(* IEC 61131-3 sources: nautilus/examples/it-cluster/lib, 2 files *)

(* ---- server.st ---- *)
(* The server half of the plant: fault inputs, a first-order thermal model,
   and how a server's parts respond. Same rules as lib/switch.st: a fault
   is an input, the recording is the baseline, faults compose, clearing a
   fault lets the recording show through again.

   The thermal model is deliberately small, and every number that shapes it
   is a named constant below, to tune against what a real box does:

     load rise    = KLoad * (CpuLoad - RecLoadPct)
     rise target  = load rise
                  + KFanFrac * failed fans * (CPU over inlet + load rise)
                  - KBoostCool * (FanBoost - 1)         the others ramping
     each sensor  = recorded + Weight * rise + room offset, approached
                    with time constant TauS (first order), so a failure
                    makes temperatures CLIMB rather than jump
     fan boost    = 1 + KBoost * (CPU rise now), capped at MaxBoost: the
                    BMC's fan curve answering the temperature it reads

   Where the numbers come from (the node is a Supermicro 1U with one
   Xeon 6505P: 150 W TDP, 97 °C DTS max; its BMC calls 102 °C critical):
     WPerPct   150 W TDP over an idle package of about 35 W, across 90 %
               of load: about 1.3 W per %
     KLoad     that power through a 1U heatsink at about 0.3 °C/W:
               about 0.35 °C per %
     KFanFrac  one of six fans gone costs the heatsink about a fifth of its
               airflow; its thermal resistance, and so the CPU's rise over
               the inlet, grows by about as much: small at idle, large
               under load, which is how a lost fan really behaves
     TauS      a 1U heatsink under forced air settles in about a minute
               (vendors give 60 s to swap a fan before cooling is lost)
     CapC      the CPU throttles near its limit rather than running away:
               held a little past the BMC's critical, so the alarm trips *)

TYPE
  SimServer : STRUCT
    Dark     : BOOL; (* the BMC stops answering: Online false *)
    PowerOff : BOOL; (* host off: standby power, fans stop, temps fall to inlet, host links drop; the BMC stays up *)
    CpuLoad  : REAL; (* % busy, 0 = as recorded (the recording is a quiet cluster, about RecLoadPct) *)
  END_STRUCT;
  SimFan : STRUCT
    Fail : BOOL; (* stopped: RPM 0, Fault; the other fans ramp, temperatures rise *)
  END_STRUCT;
  SimPSU : STRUCT
    InputLost : BOOL; (* line cord out: InputOk false, output 0, the other PSU carries the load *)
    Fail      : BOOL; (* the supply itself fails: Fault, output 0 *)
  END_STRUCT;
  SimDrive : STRUCT
    Pulled  : BOOL; (* out of its bay: Present false *)
    Failing : BOOL; (* SMART predicts failure: PredictedFailure, health Warning *)
  END_STRUCT;
  SimNetPort : STRUCT
    Down : BOOL; (* the port loses link: both ends of its cable go down *)
  END_STRUCT;
  SimCable : STRUCT
    Pulled : BOOL; (* the cable itself: both ends down *)
  END_STRUCT;
  SimRoom : STRUCT
    InletDeltaC : REAL; (* the room runs hot: every server's inlet, and everything behind it, rises *)
  END_STRUCT;
END_TYPE

FUNCTION_BLOCK ServerPlant
(* The chassis: power, CPU busy, and the thermal model's rise. Its outputs
   drive the fans, sensors and PSUs of the same server. *)
VAR_INPUT
  Rec        : Server;
  F          : SimServer;
  Room       : SimRoom;
  FansFailed : DINT;
  CpuRiseNow : REAL; (* the CPU sensor's current rise over the recording, for the fan curve *)
  CpuOverInlet : REAL := 35.0; (* the recorded CPU temperature above the recorded inlet *)
  Live       : BOOL;
  Unpowered  : BOOL; (* every supply down (plant.st): no standby power either *)
END_VAR
VAR_IN_OUT
  P : Server;
END_VAR
VAR_OUTPUT
  RiseTarget : REAL; (* °C the CPU heads for above the recording *)
  FanBoost   : REAL; (* the fans' speed factor *)
  Off        : BOOL;
  Dead       : BOOL; (* no power at all: the host off and the BMC with it *)
  LoadW      : REAL; (* the power the PSUs deliver *)
END_VAR
VAR
  B        : Server;
  Init     : BOOL;
  LoadRise : REAL;
END_VAR
VAR CONSTANT
  RecLoadPct : REAL := 10.0;  (* the recording's CPU busy: an idle cluster *)
  KLoad      : REAL := 0.35;  (* °C per % of extra load *)
  KFanFrac   : REAL := 0.2;   (* per failed fan: the share by which the CPU's rise over the inlet grows *)
  KBoost     : REAL := 0.03;  (* fan speed-up per °C of CPU rise *)
  MaxBoost   : REAL := 1.6;   (* fans at their ceiling *)
  KBoostCool : REAL := 10.0;  (* °C the ramped fans take back at full boost - 1 *)
  WPerPct    : REAL := 1.3;   (* W per % of extra load *)
  StandbyW   : REAL := 12.0;  (* host off, BMC on *)
END_VAR
IF NOT Init THEN
  B := P;
  Init := TRUE;
END_IF;
IF Live THEN
  B.PowerOn := Rec.PowerOn;
  B.PowerW := Rec.PowerW;
  B.InletTempC := Rec.InletTempC;
  B.MaxTempC := Rec.MaxTempC;
END_IF;
Dead := Unpowered;
Off := F.PowerOff OR NOT B.PowerOn OR Dead;
P.Online := NOT (F.Dark OR Dead);
P.PowerOn := NOT Off;
FanBoost := LIMIT(1.0, 1.0 + KBoost * MAX(CpuRiseNow, 0.0), MaxBoost);
IF Off THEN
  RiseTarget := 0.0;
  LoadW := SEL(Dead, StandbyW, 0.0);
  P.CpuPct := 0.0;
ELSE
  LoadRise := 0.0;
  IF F.CpuLoad > 0.0 THEN
    LoadRise := KLoad * (F.CpuLoad - RecLoadPct);
  END_IF;
  RiseTarget := LoadRise + KFanFrac * INT_TO_REAL(FansFailed) * MAX(CpuOverInlet + LoadRise, 0.0)
    - KBoostCool * (FanBoost - 1.0);
  IF F.CpuLoad > 0.0 THEN
    LoadW := B.PowerW + WPerPct * (F.CpuLoad - RecLoadPct);
    P.CpuPct := F.CpuLoad;
  ELSE
    LoadW := B.PowerW;
    P.CpuPct := RecLoadPct;
  END_IF;
END_IF;
P.PowerW := LoadW;
P.InletTempC := B.InletTempC + Room.InletDeltaC;
END_FUNCTION_BLOCK

FUNCTION_BLOCK TempPlant
(* One temperature sensor: its recording, plus Weight x the server's rise,
   plus the room; approached with TauS. Off, it cools to the inlet. *)
VAR_INPUT
  Rec        : TempSensor;
  RiseTarget : REAL;
  Weight     : REAL; (* 1 for the CPU, less for what sits further from it, 0 for the inlet *)
  RoomC      : REAL;
  InletC     : REAL; (* where it cools to, host off *)
  Off        : BOOL;
  Dt         : REAL;
  Live       : BOOL;
  CapC       : REAL := 110.0; (* where the part throttles or trips; the CPU's is lower *)
END_VAR
VAR_IN_OUT
  P : TempSensor;
END_VAR
VAR_OUTPUT
  Rise : REAL; (* now, over the recording *)
  Base : REAL; (* the recording (or snapshot) *)
END_VAR
VAR
  B     : TempSensor;
  Init  : BOOL;
  State : REAL; (* the sensor's own lagged offset from the recording *)
  Goal  : REAL;
END_VAR
VAR CONSTANT
  TauS    : REAL := 60.0;  (* heating and cooling time constant *)
  OffTauS : REAL := 300.0; (* cooling to the inlet, host off *)
END_VAR
IF NOT Init THEN
  B := P;
  Init := TRUE;
END_IF;
IF Live THEN
  B.Value := Rec.Value;
END_IF;
IF Off THEN
  Goal := InletC - B.Value;
  State := State + (Goal - State) * MIN(Dt / OffTauS, 1.0);
ELSE
  Goal := Weight * RiseTarget + RoomC;
  State := State + (Goal - State) * MIN(Dt / TauS, 1.0);
END_IF;
P.Value := MIN(B.Value + State, CapC);
Rise := P.Value - B.Value;
Base := B.Value;
P.High := P.HighSP > 0.0 AND P.Value >= P.HighSP;
P.HighHigh := P.HighHighSP > 0.0 AND P.Value >= P.HighHighSP;
END_FUNCTION_BLOCK

FUNCTION_BLOCK FanPlant
VAR_INPUT
  Rec   : Fan;
  F     : SimFan;
  Boost : REAL;
  Off   : BOOL;
  Live  : BOOL;
END_VAR
VAR_IN_OUT
  P : Fan;
END_VAR
VAR
  B    : Fan;
  Init : BOOL;
END_VAR
VAR CONSTANT
  MaxRPM : REAL := 16000.0;
END_VAR
IF NOT Init THEN
  B := P;
  Init := TRUE;
END_IF;
IF Live THEN
  B.RPM := Rec.RPM;
END_IF;
IF F.Fail OR Off THEN
  P.RPM := 0.0;
ELSE
  P.RPM := MIN(B.RPM * Boost, MaxRPM);
END_IF;
P.Fault := F.Fail;
END_FUNCTION_BLOCK

FUNCTION_BLOCK PsuPair
(* Two supplies sharing a load: each carries its recorded share while both
   are up; one lost, the other carries it all and the server stays up; both
   lost, neither carries anything (the server is Unpowered, plant.st). *)
VAR_INPUT
  Rec1, Rec2 : PSU;
  F1, F2     : SimPSU;
  LoadW      : REAL;
  Live       : BOOL;
END_VAR
VAR_IN_OUT
  P1, P2 : PSU;
END_VAR
VAR
  B1, B2 : PSU;
  Init   : BOOL;
  Up1, Up2 : BOOL;
  Share1 : REAL;
END_VAR
IF NOT Init THEN
  B1 := P1;
  B2 := P2;
  Init := TRUE;
END_IF;
IF Live THEN
  B1.InputV := Rec1.InputV;
  B1.OutputW := Rec1.OutputW;
  B2.InputV := Rec2.InputV;
  B2.OutputW := Rec2.OutputW;
END_IF;
Up1 := NOT (F1.InputLost OR F1.Fail);
Up2 := NOT (F2.InputLost OR F2.Fail);
Share1 := 0.5;
IF B1.OutputW + B2.OutputW > 0.0 THEN
  Share1 := B1.OutputW / (B1.OutputW + B2.OutputW);
END_IF;
IF NOT Up2 THEN
  Share1 := 1.0;
ELSIF NOT Up1 THEN
  Share1 := 0.0;
END_IF;
P1.OutputW := LoadW * Share1;
P2.OutputW := LoadW * (1.0 - Share1);
IF NOT (Up1 OR Up2) THEN
  P1.OutputW := 0.0;
  P2.OutputW := 0.0;
END_IF;
P1.InputOk := NOT F1.InputLost;
P2.InputOk := NOT F2.InputLost;
P1.InputV := SEL(F1.InputLost, B1.InputV, 0.0);
P2.InputV := SEL(F2.InputLost, B2.InputV, 0.0);
(* a supply with no input reports itself unhealthy, as a real one does *)
P1.Fault := NOT Up1;
P2.Fault := NOT Up2;
END_FUNCTION_BLOCK

FUNCTION_BLOCK PsuSingle
(* One supply: it carries the whole load while it is up; lost, the server
   is Unpowered (plant.st). *)
VAR_INPUT
  Rec   : PSU;
  F     : SimPSU;
  LoadW : REAL;
  Live  : BOOL;
END_VAR
VAR_IN_OUT
  P : PSU;
END_VAR
VAR
  B    : PSU;
  Init : BOOL;
  Up   : BOOL;
END_VAR
IF NOT Init THEN
  B := P;
  Init := TRUE;
END_IF;
IF Live THEN
  B.InputV := Rec.InputV;
END_IF;
Up := NOT (F.InputLost OR F.Fail);
P.OutputW := SEL(Up, 0.0, LoadW);
P.InputOk := NOT F.InputLost;
P.InputV := SEL(F.InputLost, B.InputV, 0.0);
P.Fault := NOT Up;
END_FUNCTION_BLOCK

FUNCTION_BLOCK PsuUnit
(* One of N supplies (three or more; one and two have PsuSingle and
   PsuPair). The server's draw is shared equally across the supplies that
   are up: each carries LoadW / UpCount, a supply that is down carries 0,
   and with every supply down nobody carries anything (the server is
   Unpowered, plant.st). UpCount is the number of supplies up, counted by
   plant.st from the same fault inputs in the same scan, before any unit
   runs, so a supply failing moves the share to the others in that scan,
   not the next. Each unit's own Up is the same test the count uses. *)
VAR_INPUT
  Rec     : PSU;
  F       : SimPSU;
  LoadW   : REAL;
  UpCount : DINT; (* supplies up on this server, this scan *)
  Live    : BOOL;
END_VAR
VAR_IN_OUT
  P : PSU;
END_VAR
VAR
  B    : PSU;
  Init : BOOL;
  Up   : BOOL;
END_VAR
IF NOT Init THEN
  B := P;
  Init := TRUE;
END_IF;
IF Live THEN
  B.InputV := Rec.InputV;
END_IF;
Up := NOT (F.InputLost OR F.Fail);
P.OutputW := SEL(Up AND UpCount > 0, 0.0, LoadW / INT_TO_REAL(MAX(UpCount, 1)));
P.InputOk := NOT F.InputLost;
P.InputV := SEL(F.InputLost, B.InputV, 0.0);
P.Fault := NOT Up;
END_FUNCTION_BLOCK

FUNCTION_BLOCK DrivePlant
VAR_INPUT
  F : SimDrive;
END_VAR
VAR_IN_OUT
  P : Drive;
END_VAR
P.Present := NOT F.Pulled;
P.PredictedFailure := F.Failing;
IF F.Failing THEN
  P.Health := 1;
ELSE
  P.Health := 0;
END_IF;
P.Fault := P.Health > 0 OR NOT P.Present;
END_FUNCTION_BLOCK

FUNCTION_BLOCK NicPlant
(* A server's network port. LinkOk is its cable's state, worked out once
   per cable from both ends' faults (plant.st), so a port down at the
   switch drops the server's end too: the cable goes dark at both ends. *)
VAR_INPUT
  Rec       : NetPort;
  LinkOk    : BOOL;
  SpeedGbps : REAL; (* the cable's negotiated speed override, 0 = as recorded *)
  Live      : BOOL;
END_VAR
VAR_IN_OUT
  P : NetPort;
END_VAR
VAR
  B    : NetPort;
  Init : BOOL;
END_VAR
IF NOT Init THEN
  B := P;
  Init := TRUE;
END_IF;
IF Live THEN
  B.LinkUp := Rec.LinkUp;
  B.SpeedGbps := Rec.SpeedGbps;
END_IF;
P.LinkUp := B.LinkUp AND LinkOk;
IF NOT P.LinkUp THEN
  P.SpeedGbps := 0.0;
ELSIF SpeedGbps > 0.0 THEN
  P.SpeedGbps := SpeedGbps;
ELSE
  P.SpeedGbps := B.SpeedGbps;
END_IF;
END_FUNCTION_BLOCK

(* ---- switch.st ---- *)
(* The switch half of the plant: fault inputs, and how they bend a port.

   A fault is an INPUT, never a value: the recording stays the source of
   every member no fault touches, and faults compose (a port can be
   speed-degraded AND erroring, with its switch dark over all of it).
   Clear the input and the recording shows through again. Write them from
   the HMI (Set Live Value), `curl .../api/tags`, or a test's given:. *)

TYPE
  SimPort : STRUCT
    Down      : BOOL; (* link lost: OperUp false, no traffic; admin stays up, so the monitor alarms *)
    AdminDown : BOOL; (* shut by an operator: AdminUp and OperUp false, not an alarm *)
    SpeedMbps : REAL; (* negotiated speed override, both ends of the cable, 0 = as recorded (10000 to 1000: degraded) *)
    ErrorRate : REAL; (* extra errors per second on top of the recording *)
    (* VLANs, applied in plant.st over the configured membership: *)
    Pvid      : DINT; (* native VLAN override, 0 = as configured (a native mismatch) *)
    Prune     : DINT; (* a VLAN taken off the port, 0 = none (a trunk missing a VLAN) *)
    Access    : DINT; (* the port moved to this access VLAN alone, 0 = as configured *)
  END_STRUCT;
  SimNet : STRUCT
    (* the layer-2 domain, all three switches trunked on their ring: a storm
       floods every port that has link *)
    BroadcastPps : REAL; (* a broadcast storm: packets per second flooded out of every up port *)
    MulticastPps : REAL; (* a multicast flood, the same way (no IGMP snooping to stop it) *)
  END_STRUCT;
  SimSwitch : STRUCT
    Dark   : BOOL; (* the switch stops answering: every port down, the agent silent *)
    Reboot : BOOL; (* a pulse: dark for RebootS, then back with its uptime reset; clears itself (ClearFaults ends it early) *)
  END_STRUCT;
END_TYPE

FUNCTION SlowerMbps : REAL
(* Two speed overrides on one link, 0 = none: the slower one, as the two
   ends negotiate it. *)
VAR_INPUT
  A : REAL;
  B : REAL;
END_VAR
IF A > 0.0 AND (B <= 0.0 OR A < B) THEN
  SlowerMbps := A;
ELSIF B > 0.0 THEN
  SlowerMbps := B;
ELSE
  SlowerMbps := 0.0;
END_IF;
END_FUNCTION

FUNCTION_BLOCK PortPlant
(* One switch port. P is the port as the device reports it: its identity
   (Name, Index, Alias, counters) is its own and never touched here; the
   members the recording carries follow Rec while the replay is Live, and
   hold the tag's initial snapshot while it is not (no recording loaded),
   so a plant without its data still reports a plausible, quiet switch. *)
VAR_INPUT
  Rec  : SwitchPort; (* the recording, from the replay driver *)
  F    : SimPort;    (* this port's faults *)
  Dark : BOOL;       (* the switch's *)
  Live : BOOL;       (* the recording is playing *)
  LinkOk : BOOL := TRUE; (* its cable, from both ends' faults (plant.st); TRUE unwired *)
  LinkMbps : REAL := 0.0; (* its cable's speed override, from both ends' faults (plant.st); 0 = none *)
  Net  : SimNet;     (* a storm in the layer-2 domain *)
  Dt   : REAL;       (* seconds since the last scan, for the discard counter *)
END_VAR
VAR_IN_OUT
  P : SwitchPort;
END_VAR
VAR
  B        : SwitchPort; (* the baseline: recording or snapshot, never a fault *)
  Init     : BOOL;
  FloodBps : REAL;
  LineBps  : REAL;
  Dropped  : REAL; (* discards not yet whole, so the counter never loses a fraction *)
  DropPps  : REAL; (* frames the line cannot carry, per second *)
  Mbps     : REAL; (* the speed override in force: this port's, or its cable's if slower *)
END_VAR
VAR CONSTANT
  FloodBytes : REAL := 128.0; (* a storm's frames are small: ARP, discovery, a looped packet *)
END_VAR
IF NOT Init THEN
  B := P;
  Init := TRUE;
END_IF;
IF Live THEN
  B.AdminUp := Rec.AdminUp;
  B.OperUp := Rec.OperUp;
  B.SpeedMbps := Rec.SpeedMbps;
  B.InBps := Rec.InBps;
  B.OutBps := Rec.OutBps;
  B.ErrorRate := Rec.ErrorRate;
END_IF;
P.AdminUp := B.AdminUp AND NOT F.AdminDown;
P.OperUp := B.OperUp AND LinkOk AND NOT (F.Down OR F.AdminDown OR Dark);
P.SpeedMbps := B.SpeedMbps;
P.InBps := B.InBps;
P.OutBps := B.OutBps;
(* a link runs at one speed: an override at either end of the cable is
   this end's too *)
Mbps := SlowerMbps(A := F.SpeedMbps, B := LinkMbps);
IF Mbps > 0.0 AND P.OperUp THEN
  P.SpeedMbps := Mbps;
  (* traffic cannot exceed the line *)
  P.InBps := MIN(P.InBps, Mbps * 1000000.0);
  P.OutBps := MIN(P.OutBps, Mbps * 1000000.0);
END_IF;
DropPps := 0.0;
IF NOT P.OperUp THEN
  P.InBps := 0.0;
  P.OutBps := 0.0;
  P.InBroadcastPps := 0.0;
  P.InMulticastPps := 0.0;
ELSE
  (* a storm: every up port receives the flood and sends it on; what the
     line cannot carry is dropped, and counted *)
  P.InBroadcastPps := B.InBroadcastPps + Net.BroadcastPps;
  P.InMulticastPps := B.InMulticastPps + Net.MulticastPps;
  FloodBps := (Net.BroadcastPps + Net.MulticastPps) * FloodBytes * 8.0;
  LineBps := P.SpeedMbps * 1000000.0;
  P.InBps := MIN(P.InBps + FloodBps, LineBps);
  P.OutBps := P.OutBps + FloodBps;
  IF LineBps > 0.0 AND P.OutBps > LineBps THEN
    DropPps := (P.OutBps - LineBps) / (FloodBytes * 8.0);
    Dropped := Dropped + DropPps * Dt;
    P.OutBps := LineBps;
  END_IF;
  IF Dropped >= 1.0 THEN
    P.OutDiscards := P.OutDiscards + REAL_TO_INT(Dropped - 0.5);
    Dropped := Dropped - INT_TO_REAL(REAL_TO_INT(Dropped - 0.5));
  END_IF;
END_IF;
P.ErrorRate := B.ErrorRate + F.ErrorRate;
P.DiscardRate := DropPps; (* the stand-in integrates ifOutDiscards from it *)
P.Down := P.AdminUp AND NOT P.OperUp;
IF P.SpeedMbps > 0.0 THEN
  P.InPct := 100.0 * P.InBps / (P.SpeedMbps * 1000000.0);
  P.OutPct := 100.0 * P.OutBps / (P.SpeedMbps * 1000000.0);
ELSE
  P.InPct := 0.0;
  P.OutPct := 0.0;
END_IF;
END_FUNCTION_BLOCK

FUNCTION_BLOCK SwitchPlant
(* The chassis: dark, rebooting, and its uptime, which counts while it is
   up and starts again from 0 after a reboot. *)
VAR_INPUT
  Dt    : REAL;
  Clear : BOOL; (* ClearFaults this scan: a reboot in progress ends *)
END_VAR
VAR_IN_OUT
  F : SimSwitch;
  P : Switch;
END_VAR
VAR_OUTPUT
  Down : BOOL; (* dark or rebooting: its ports and their cables are down *)
END_VAR
VAR
  T         : TON;
  Rebooting : BOOL;
  Up        : REAL;
  Init      : BOOL;
END_VAR
VAR CONSTANT
  RebootS : TIME := T#90S;
END_VAR
IF NOT Init THEN
  Up := INT_TO_REAL(P.UptimeS);
  Init := TRUE;
END_IF;
IF F.Reboot THEN
  Rebooting := TRUE;
  F.Reboot := FALSE;
END_IF;
IF Clear THEN
  Rebooting := FALSE;
END_IF;
T(IN := Rebooting, PT := RebootS);
IF T.Q THEN
  Rebooting := FALSE;
  Up := 0.0;
END_IF;
Down := F.Dark OR Rebooting;
IF NOT Down THEN
  Up := Up + Dt;
END_IF;
P.Online := NOT Down;
P.UptimeS := REAL_TO_INT(Up);
END_FUNCTION_BLOCK
